FUNCTION Celsius_To_Farenheit : REAL
VAR_INPUT
	fCelsius : REAL;
END_VAR
VAR
END_VAR

Celsius_To_Farenheit := fCelsius * 1.8 + 32;

END_FUNCTION

(* stored: Version 1.1.0.1
   POU Celsius_To_Farenheit: Id {7920b028-4bc7-41f6-b576-dff1b341345d}, SpecialFunc None *)
